// TIA Portal V20 export
// export: Created 2026-10-19T18:04:23.843683Z, ExportSetting WithDefaults, DisplayName Totally Integrated Automation Portal, DisplayVersion V20 Update 6, DisplayName TIA Portal Openness, DisplayVersion V20 Update 6, DisplayName TIA Portal Version Control Interface, DisplayVersion V20 Update 6, DisplayName SINAMICS Startdrive Advanced, DisplayVersion V20 SP1, DisplayName SINAMICS Startdrive G130, G150, S120, S150, SINAMICS MV, G220, S200, S210, DisplayVersion V20 SP1, DisplayName SINAMICS Startdrive G110M, G120, G120C, G120D, G120P, G115D, DisplayVersion V20 SP1, DisplayName STEP 7 Professional, DisplayVersion V20 Update 6, DisplayName STEP 7 Safety, DisplayVersion V20 Update 2, DisplayName WinCC Basic/Comfort/Advanced, DisplayVersion V20 Update 6, DisplayName WinCC Unified, DisplayVersion V20 Update 6
FUNCTION "GeneralErros_HMII" : Void   // FC13, SCL
{ S7_Optimized_Access := 'TRUE' }
VERSION : 0.1
// stored: AutoNumber true, IsIECCheckEnabled false, SetENOAutomatically false, UDAEnableTagReadback false
BEGIN
   "HMI_DB".GeneralErrors.%X0 := "Control_DB".LCnv_Control[1].Safety_Stop_Cnrl.Error;
   "HMI_DB".GeneralErrors.%X1 := "Control_DB".LCnv_Control[1].Safety_Stop_Cnrl.Error;
   "HMI_DB".GeneralErrors.%X2 := "Control_DB".LCnv_Control[2].Safety_Stop_Cnrl.Error;
   "HMI_DB".GeneralErrors.%X3 := "Control_DB".LCnv_Control[2].Safety_Stop_Cnrl.Error;
   "HMI_DB".GeneralErrors.%X4 := "Control_DB".LCnv_Control[3].Safety_Stop_Cnrl.Error;
   "HMI_DB".GeneralErrors.%X5 := "Control_DB".LCnv_Control[3].Safety_Stop_Cnrl.Error;

   "Error" := "System_DB_VTD".Error OR "System_DB_Carousel".Error;
END_FUNCTION
